RoboDK station: kuka_station.rdk

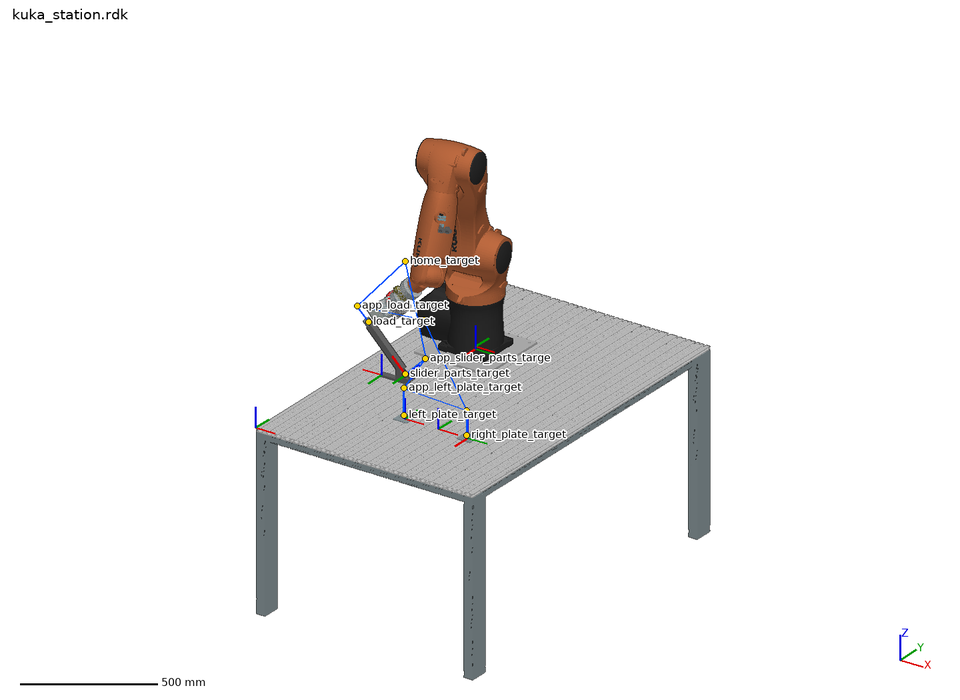
[picture v0: the station drawn from its stored meshes, robots at their saved joint values, targets as dots, program paths as lines]
Station kuka_station (saved by RoboDK 6.0.7). Poses are relative to the parent item; angles as X-Y-Z fixed-axis rotations.
  - frame table_frame at (0, 0, 0) mm
    - object table_object at (0, 0, 0) mm, size 960.1 x 1500 x 750 mm, geometry from table_object.sld
    - target home_target (Cartesian target) at (280, 545, 532) mm, rotated rx 180 ry 0 rz 47 deg; joints [90, -90, 90, 0, 90, 0] of KUKA KR 6 R900 sixx
    - target left_plate_target (Cartesian target) at (396, 370, 13) mm, rotated rx -180 ry 0 rz 0 deg; joints [79.403, -41.229, 97.284, 0, 33.945, -57.597] of KUKA KR 6 R900 sixx
    - target app_left_plate_target (Cartesian target) at (396, 370, 123) mm, rotated rx -180 ry 0 rz 0 deg; joints [79.403, -51.193, 96.429, 0, 44.764, -57.597] of KUKA KR 6 R900 sixx
    - target right_plate_target (Cartesian target) at (677.82, 366.9, 12.54) mm, rotated rx -180 ry 0 rz -88.78 deg; joints [57.444, -31.46, 75.522, 0, 45.939, -168.336] of KUKA KR 6 R900 sixx
    - target app_right_plate_target (Cartesian target) at (677.82, 366.9, 112.54) mm, rotated rx -180 ry 0 rz -88.78 deg; joints [57.444, -39.155, 74.87, 0, 54.285, -168.336] of KUKA KR 6 R900 sixx
    - target slider_parts_target (Cartesian target) at (230.58, 617, 34.24) mm, rotated rx 180 ry 45 rz 0 deg; joints [60.528, -41.46, 127.701, 57.413, 46.939, -132.52] of KUKA KR 6 R900 sixx
    - target app_slider_parts_target (Cartesian target) at (318.97, 617, 122.62) mm, rotated rx -180 ry 45 rz 0 deg; joints [51.267, -51.817, 122.511, 40.26, 58.596, -119.412] of KUKA KR 6 R900 sixx
    - target load_target (Cartesian target) at (63.91, 620.52, 197.08) mm, rotated rx 180 ry 45 rz 0 deg; joints [83.189, -69.258, 137.839, 64.407, 51.123, -109.239] of KUKA KR 6 R900 sixx
    - target app_load_target (Cartesian target) at (14.42, 620.52, 246.58) mm, rotated rx -180 ry 45 rz 0 deg; joints [90.832, -76.777, 136.755, 63.997, 51.875, -97.51] of KUKA KR 6 R900 sixx
    - frame base_plate_frame at (280, 990, 0) mm, rotated rx 0 ry 0 rz -90 deg
      - object base_plate_object at (0, 0, 0) mm, size 320 x 320 x 10 mm, geometry from base_plate_object.sld
    - frame slider_frame at (125, 617, 0) mm, rotated rx 0 ry 0 rz 180 deg
      - object slider_object at (0, 0, 0) mm, size 198.7 x 26 x 198.7 mm, 1 curves, geometry from slider_object.sld
    - frame slider_parts_frame at (232.7, 617, 30.7) mm, rotated rx 0 ry -45 rz -180 deg
    - frame pick_and_drop_frame at (550, 370, 0) mm
    - frame right_frame at (680, 370, 0) mm, rotated rx 0 ry 0 rz -90 deg
      - object right_plate_object at (0, 0, 0) mm, size 60 x 60 x 9 mm, 1 curves, geometry from right_plate_object.sld
    - frame left_frame at (400, 370, 0) mm
      - object left_plate_object at (0, 0, 0) mm, size 60 x 60 x 9 mm, 1 curves, geometry from left_plate_object.sld
    - frame kuka_frame at (280, 990, 10) mm
      - robot KUKA KR 6 R900 sixx: 6 axes, payload 6 kg, reach 901 mm, repeatability 0.03 mm, weight 52 kg
          modified DH rows (alpha deg, a mm, theta deg, d mm): 0, 0, 0, 400; -90, 25, 0, 0; 0, 455, -90, 0; -90, 35, 0, 420; 90, 0, 0, 0; -90, 0, 180, 80
          joint limits [-170, -190, -120, -185, -120, -350] to [170, 45, 156, 185, 120, 350]; home [0, -90, 90, 0, 0, 0]; saved at [83.189, -69.258, 137.839, 64.407, 51.123, -109.239]
        - tool gripper_TCP, TCP at (0, 0, 288) mm, rotated rx 0 ry 0 rz 43 deg
        - robot gripper: 1 axes
            joint limits [0] to [50]; home [0]; saved at [50]
    - target close_gripper_target (joint target) at (-24.9, 610.96, 271.99) mm, rotated rx -174.53 ry 42.03 rz 5.46 deg; joints [20, -78.968, 131.593, 59.422, 51.098, -80.049] of gripper
    - target open_gripper_target (joint target) at (-24.9, 610.96, 271.99) mm, rotated rx -174.53 ry 42.03 rz 5.46 deg; joints [50, -78.968, 131.593, 59.422, 51.098, -80.049] of gripper
    - target pre_app_load_target (Cartesian target) at (322.68, 604.39, 282.54) mm, rotated rx -180 ry 0 rz -88.78 deg; joints [83.684, -89.981, 125.332, 0, 54.649, -142.096] of KUKA KR 6 R900 sixx
    - object part_object at (65.6, 620.52, 192.54) mm, rotated rx 0 ry -45 rz 180 deg, size 40 x 20 x 20 mm, 1 curves, geometry from part_object.sld
  - folder programs
    - program factory_reset (1 instructions, listed below)
    - program open_gripper (3 instructions, listed below)
    - program close_gripper (3 instructions, listed below)
    - program main (35 instructions, listed below)
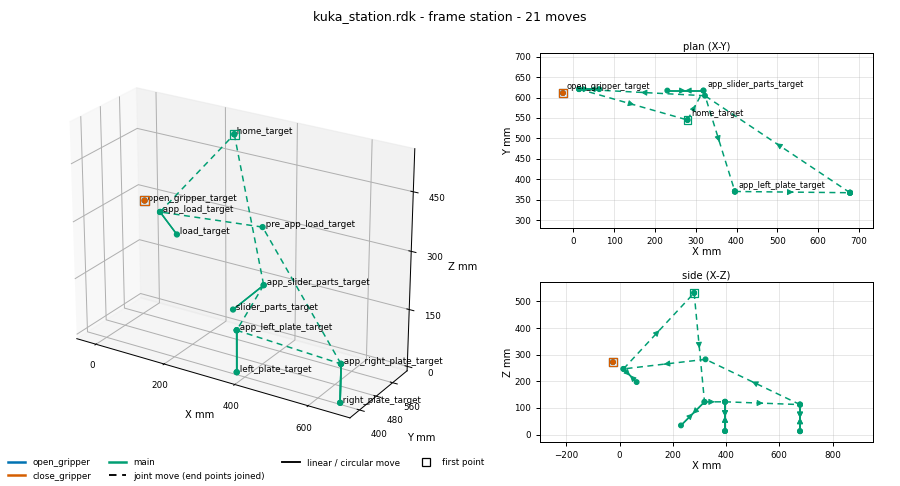
[picture p0: tool path of kuka_station.rdk in frame station, 21 of 21 moves have a stored position in this frame; points joined in program order, loops and branches not executed]

--- program factory_reset (robot KUKA KR 6 R900 sixx) ---
  Move objects

--- program open_gripper (robot gripper) ---
  Set Ref.: table_frame
  Set Tool: gripper_TCP
  MoveJ (open_gripper_target)

--- program close_gripper (robot gripper) ---
  Set Ref.: table_frame
  Set Tool: gripper_TCP
  MoveJ (close_gripper_target)

--- program main (robot KUKA KR 6 R900 sixx) ---
  Call factory_reset
  Set Ref.: table_frame
  Set Tool: gripper_TCP
  MoveJ (home_target)
  Call open_gripper
  MoveJ (app_slider_parts_target)
  MoveL (slider_parts_target)
  Call close_gripper
  Attach to gripper_TCP
  MoveL (app_slider_parts_target)
  MoveJ (app_left_plate_target)
  MoveL (left_plate_target)
  Call open_gripper
  Detach from gripper_TCP
  MoveL (app_left_plate_target)
  MoveL (left_plate_target)
  Call close_gripper
  Attach to gripper_TCP
  MoveL (app_left_plate_target)
  MoveJ (app_right_plate_target)
  MoveL (right_plate_target)
  Call open_gripper
  Detach from gripper_TCP
  MoveL (app_right_plate_target)
  MoveL (right_plate_target)
  Call close_gripper
  Attach to gripper_TCP
  MoveL (app_right_plate_target)
  MoveJ (pre_app_load_target)
  MoveJ (app_load_target)
  MoveL (load_target)
  Call open_gripper
  Detach from gripper_TCP
  MoveL (app_load_target)
  MoveJ (home_target)
